(* IEC 61131-3 sources: trust-platform/crates/trust-runtime/tests/fixtures/ci/broken/src, 1 file *)

(* ---- main.st ---- *)
PROGRAM Main
VAR
    Count : INT := 0;
END_VAR

Count := Count + 1;
END_PROGRAM
